(* IEC 61131-3 sources: llm-plc-st-eval/data/processed_definitivo/qwen2.5-coder_14b/B7/few_shot, 3 files *)

(* ---- ejec_1.st ---- *)
FUNCTION_BLOCK SelBomba
VAR_INPUT
    modoAuto : BOOL; (* Modo automático *)
    btnManual : BOOL; (* Botón manual *)
    nivelBajo : BOOL; (* Nivel bajo *)
END_VAR
VAR_OUTPUT
    bomba : BOOL; (* Estado de la bomba *)
END_VAR

(* Selección de la fuente de mando *)
IF modoAuto THEN
    bomba := nivelBajo; (* En modo automático, la bomba está encendida si el nivel está bajo *)
ELSE
    bomba := btnManual; (* En modo manual, la bomba obedece al botón manual *)
END_IF
END_FUNCTION_BLOCK

(* ---- ejec_2.st ---- *)
FUNCTION_BLOCK SelBomba
VAR_INPUT
    modoAuto : BOOL; (* Modo automático *)
    btnManual : BOOL; (* Botón manual *)
    nivelBajo : BOOL; (* Nivel bajo *)
END_VAR
VAR_OUTPUT
    bomba : BOOL; (* Estado de la bomba *)
END_VAR

(* Selección de la fuente de mando de la bomba *)
IF modoAuto THEN
    bomba := nivelBajo; (* En modo automático, la bomba está encendida si el nivel está bajo *)
ELSE
    bomba := btnManual; (* En modo manual, la bomba obedece al botón manual *)
END_IF
END_FUNCTION_BLOCK

(* ---- ejec_3.st ---- *)
FUNCTION_BLOCK SelBomba
VAR_INPUT
    modoAuto : BOOL; (* Modo automático *)
    btnManual : BOOL; (* Botón manual *)
    nivelBajo : BOOL; (* Nivel bajo *)
END_VAR
VAR_OUTPUT
    bomba : BOOL; (* Estado de la bomba *)
END_VAR

(* Selección de la fuente de mando de la bomba *)
IF modoAuto THEN
    bomba := nivelBajo; (* En modo automático, la bomba está encendida si el nivel está bajo *)
ELSE
    bomba := btnManual; (* En modo manual, la bomba obedece al botón manual *)
END_IF
END_FUNCTION_BLOCK
